// FB TON state codes.
{attribute 'qualified_only'}
{attribute 'to_string'}
TYPE
E_SafeTonState :
(
    Undefined := 0,
    Run := 1,
    Stop := 2,
    Safe := 3,
    DelayIn := 9
) BYTE;
END_TYPE

(* stored: Version 1.1.0.1
   DUT E_SafeTonState: Id {ca8dc299-734f-5408-9a6b-64869f835c52} *)
